// TIA Portal project "PROYECTO_FINALll" (V19)

(* hardware
DEVICE "PC-System_2"  SIMATIC PC station
   slot 0: "PC station"  Rail  SIMATIC PC-Station  V1.0
      slot 125: "Stationmanager"  Station_Manager  V6.0.4
   slot 1: "HMI_RT_1"  WinCC RT Advanced  6AV2 104-0xxxx-xxxx  17.0.0.0
      slot 33792: "Computer interface"  Host interface
   slot 2: "IE general_1"  IE General  IE_CP  V8.2.0
      slot 1: "PROFINET interface"  IEGeneral.Interface.8.2.0
DEVICE "S7-1200 station_2"  S7-1200 Station
   slot 0: "Rack_0"  S7-1200 Rack  Rack  V1.0
   slot 1: "PLC_2"  CPU 1212C AC/DC/Rly  6ES7 212-1BE40-0XB0  V4.5
   slot 101: "CM 1243-5"  CM 1243-5  6GK7 243-5DX30-0XE0  V1.3
DEVICE "GSD device_1"  GSD.Device
   slot 0: "Rack_0"  Rail
*)

// ===== PLC "PLC_2"  CPU 1212C AC/DC/Rly =====

VAR_GLOBAL   // PLC tag table "Default tag table"
   "Tag_1" AT %IW68 : Int;
   "Tag_2" AT %IW70 : Int;
   "Tag_3" AT %IW72 : Word;
   "Tag_4" AT %IW74 : Int;
   "Tag_5" AT %IW76 : Int;
   "Tag_6" AT %IW78 : Int;
END_VAR

DATA_BLOCK "Data"   // DB1
{ S7_Optimized_Access := 'TRUE' }
VERSION : 0.1
   VAR
      TEMP_A : Real;
      TEMP_M : Real;
      IRRADIANCIA : Real;
      SOILING : Real;
      VOLT_MED : Real;
      CORRIENTE_MED : Real;
      VDC : Real;
      IDC : Real;
      PAC : Real;
      PR : Real;
      YF : Real;
      EAC : Real;
      PERD_SUCIEDAD : Real;
      PERD_TEMP : Real;
      "ON/OFF" : Bool;
      DEFAULT : Bool;
   END_VAR
BEGIN
END_DATA_BLOCK

DATA_BLOCK "V_AMBIENTALES_DB"   // DB2
{ S7_Optimized_Access := 'TRUE' }
VERSION : 0.1
// stored: InstanceOfName V_AMBIENTALES
"V_AMBIENTALES"
BEGIN
END_DATA_BLOCK

DATA_BLOCK "Block_1_DB"   // DB3
{ S7_Optimized_Access := 'TRUE' }
VERSION : 0.1
// stored: InstanceOfName Block_1
"Block_1"
BEGIN
END_DATA_BLOCK

DATA_BLOCK "Block_1_DB_1"   // DB4
{ S7_Optimized_Access := 'TRUE' }
VERSION : 0.1
// stored: InstanceOfName Block_1
"Block_1"
BEGIN
END_DATA_BLOCK

FUNCTION_BLOCK "V_AMBIENTALES"   // FB1, LAD
{ S7_Optimized_Access := 'TRUE' }
VERSION : 0.1
   VAR_OUTPUT
      TEMP_M : Real;
      TEMP_A : Real;
      IRRADIANCIA : Real;
      SUCIEDAD : Real;
      VOLTAJE : Real;
      CORRIENTE : Real;
   END_VAR
   VAR_TEMP
      Temp_1 : Real;
      Temp_2 : Real;
      Temp_3 : Real;
      Temp_4 : Real;
      Temp_5 : Real;
      Temp_6 : Real;
   END_VAR
BEGIN

REGION Network 1: TEMPERATURA DEL MODULO
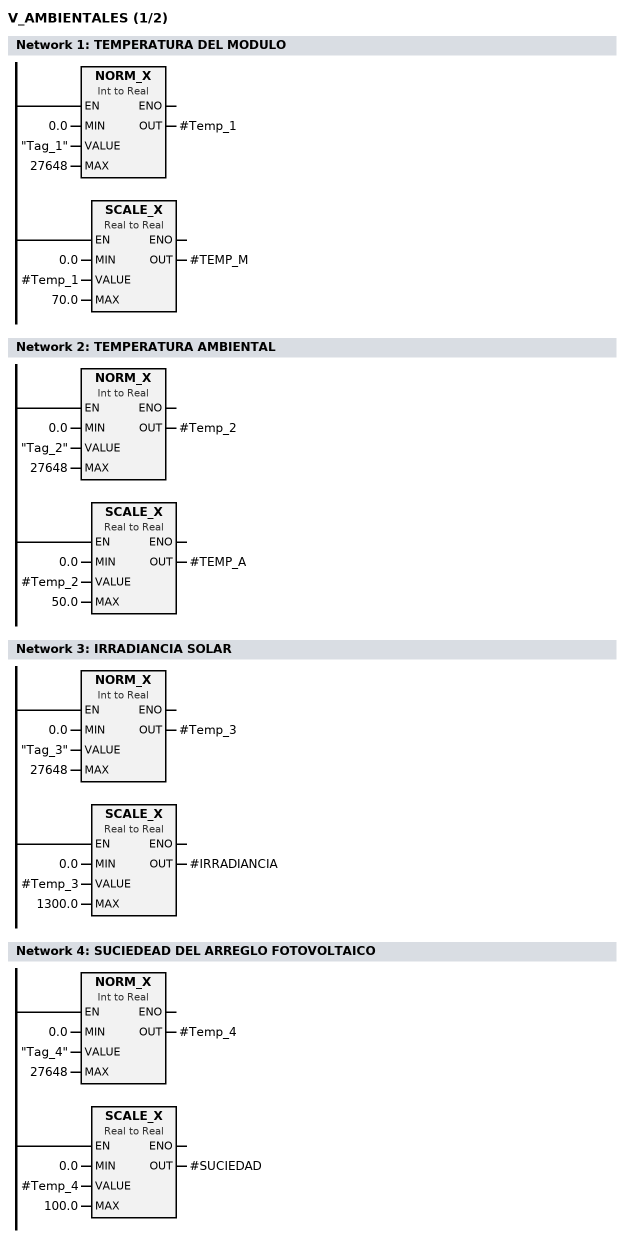
   RUNG wire#powerrail
      { S7_Templates := "[SrcType := Int, DestType := Real]" } Normalize(min := 0.0, value := "Tag_1", max := 27648, out => #Temp_1)
   END_RUNG
   RUNG wire#powerrail
      { S7_Templates := "[SrcType := Real, DestType := Real]" } Scale(min := 0.0, value := #Temp_1, max := 70.0, out => #TEMP_M)
   END_RUNG
   // the same network as SCL:
   #Temp_1 := NORM_X(MIN := 0.0, VALUE := "Tag_1", MAX := 27648);
   #TEMP_M := SCALE_X(MIN := 0.0, VALUE := #Temp_1, MAX := 70.0);
END_REGION

REGION Network 2: TEMPERATURA AMBIENTAL
   RUNG wire#powerrail
      { S7_Templates := "[SrcType := Int, DestType := Real]" } Normalize(min := 0.0, value := "Tag_2", max := 27648, out => #Temp_2)
   END_RUNG
   RUNG wire#powerrail
      { S7_Templates := "[SrcType := Real, DestType := Real]" } Scale(min := 0.0, value := #Temp_2, max := 50.0, out => #TEMP_A)
   END_RUNG
   // the same network as SCL:
   #Temp_2 := NORM_X(MIN := 0.0, VALUE := "Tag_2", MAX := 27648);
   #TEMP_A := SCALE_X(MIN := 0.0, VALUE := #Temp_2, MAX := 50.0);
END_REGION

REGION Network 3: IRRADIANCIA SOLAR
   RUNG wire#powerrail
      { S7_Templates := "[SrcType := Int, DestType := Real]" } Normalize(min := 0.0, value := "Tag_3", max := 27648, out => #Temp_3)
   END_RUNG
   RUNG wire#powerrail
      { S7_Templates := "[SrcType := Real, DestType := Real]" } Scale(min := 0.0, value := #Temp_3, max := 1300.0, out => #IRRADIANCIA)
   END_RUNG
   // the same network as SCL:
   #Temp_3 := NORM_X(MIN := 0.0, VALUE := "Tag_3", MAX := 27648);
   #IRRADIANCIA := SCALE_X(MIN := 0.0, VALUE := #Temp_3, MAX := 1300.0);
END_REGION

REGION Network 4: SUCIEDEAD DEL ARREGLO FOTOVOLTAICO
   RUNG wire#powerrail
      { S7_Templates := "[SrcType := Int, DestType := Real]" } Normalize(min := 0.0, value := "Tag_4", max := 27648, out => #Temp_4)
   END_RUNG
   RUNG wire#powerrail
      { S7_Templates := "[SrcType := Real, DestType := Real]" } Scale(min := 0.0, value := #Temp_4, max := 100.0, out => #SUCIEDAD)
   END_RUNG
   // the same network as SCL:
   #Temp_4 := NORM_X(MIN := 0.0, VALUE := "Tag_4", MAX := 27648);
   #SUCIEDAD := SCALE_X(MIN := 0.0, VALUE := #Temp_4, MAX := 100.0);
END_REGION

REGION Network 5: VOLTAJE DC
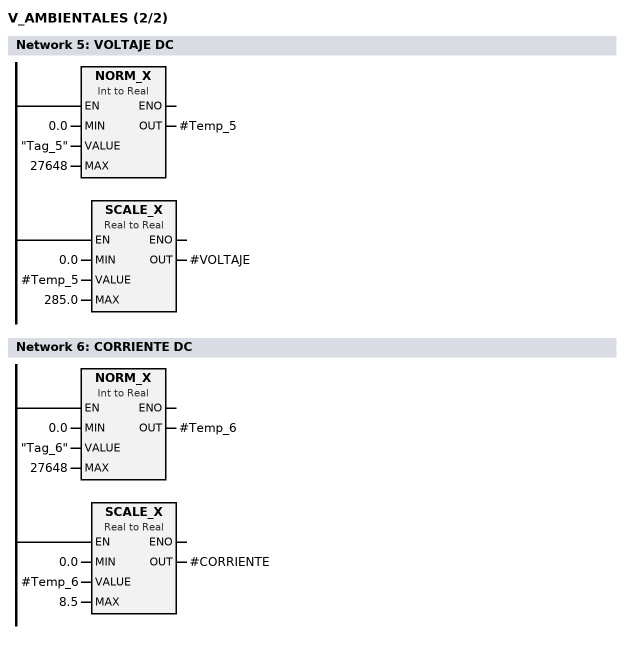
   RUNG wire#powerrail
      { S7_Templates := "[SrcType := Int, DestType := Real]" } Normalize(min := 0.0, value := "Tag_5", max := 27648, out => #Temp_5)
   END_RUNG
   RUNG wire#powerrail
      { S7_Templates := "[SrcType := Real, DestType := Real]" } Scale(min := 0.0, value := #Temp_5, max := 285.0, out => #VOLTAJE)
   END_RUNG
   // the same network as SCL:
   #Temp_5 := NORM_X(MIN := 0.0, VALUE := "Tag_5", MAX := 27648);
   #VOLTAJE := SCALE_X(MIN := 0.0, VALUE := #Temp_5, MAX := 285.0);
END_REGION

REGION Network 6: CORRIENTE DC
   RUNG wire#powerrail
      { S7_Templates := "[SrcType := Int, DestType := Real]" } Normalize(min := 0.0, value := "Tag_6", max := 27648, out => #Temp_6)
   END_RUNG
   RUNG wire#powerrail
      { S7_Templates := "[SrcType := Real, DestType := Real]" } Scale(min := 0.0, value := #Temp_6, max := 8.5, out => #CORRIENTE)
   END_RUNG
   // the same network as SCL:
   #Temp_6 := NORM_X(MIN := 0.0, VALUE := "Tag_6", MAX := 27648);
   #CORRIENTE := SCALE_X(MIN := 0.0, VALUE := #Temp_6, MAX := 8.5);
END_REGION
END_FUNCTION_BLOCK

FUNCTION_BLOCK "CALCULOS"   // FB2, LAD
{ S7_Optimized_Access := 'TRUE' }
VERSION : 0.1
   VAR_OUTPUT
      VOLTAJE_DC : Real;
   END_VAR
   VAR_TEMP
      TEMP_1 : Real;
      TEMP_2 : Real;
   END_VAR
BEGIN

REGION Network 1
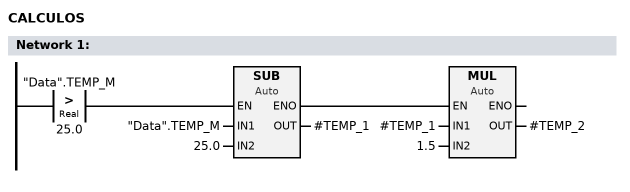
   RUNG wire#powerrail
      { S7_Templates := "SrcType := Real" } GT_Contact(in1 := "Data".TEMP_M, in2 := 25.0)
      Sub(in1 := "Data".TEMP_M, in2 := 25.0, out => #TEMP_1)
      Mul(in1 := #TEMP_1, in2 := 1.5, out => #TEMP_2)
   END_RUNG
   // the same network as SCL:
   IF "Data".TEMP_M > 25.0 THEN
       #TEMP_1 := "Data".TEMP_M - 25.0;
       #TEMP_2 := #TEMP_1 * 1.5;
   END_IF;
END_REGION
END_FUNCTION_BLOCK

FUNCTION_BLOCK "Block_1"   // FB3, SCL
{ S7_Optimized_Access := 'TRUE' }
VERSION : 0.1
   VAR_INPUT
      G_POA : Real;
      Tmod : Real;
      SR : Real;
      dt_s : Real;
      Enable : Bool;
      ResetDaily : Bool;
   END_VAR
   VAR_OUTPUT
      Vdc : Real;
      Idc : Real;
      Pac : Real;
      Eac : Real;
      Hpoa : Real;
      PR : Real;
      Yf : Real;
      Loss_soil : Real;
      Loss_therm : Real;
   END_VAR
   VAR
      P0_kw : Real := 2.25;
      Vdc_ref : Real := 282.0;
      Pac_max : Real := 2.0;
      eta_inv : Real := 0.96;
      gammaP : Real := 0.004;
      betaV : Real := 0.0035;
   END_VAR
   VAR_TEMP
      Geff : Real;
      Pdc : Real;
      tempFacP : Real;
      tempFacV : Real;
   END_VAR
BEGIN



   // Reset diario (por botón o por reloj)
   IF #ResetDaily THEN
       #Eac := 0.0;
       #Hpoa := 0.0;
   END_IF;

   IF NOT #Enable THEN
       // Si está deshabilitado, puedes congelar o poner en cero
       #Pac := 0.0;
       #Idc := 0.0;
       // Vdc lo puedes mantener o llevar a 0
       // Vdc := 0.0;
       #PR := 0.0;
       #Yf := #Eac / #P0_kw; // opcional
       RETURN;
   END_IF;

   // ---- Normalización y límites de SR ----
   // Si SR viene como porcentaje (0..100), lo convertimos a 0..1
   IF #SR > 1.5 THEN
       #SR := #SR / 100.0;
   END_IF;

   // Limitar SR a 0..1
   IF #SR < 0.0 THEN
       #SR := 0.0;
   ELSIF #SR > 1.0 THEN
       #SR := 1.0;
   END_IF;

   // ---- Pérdida por suciedad (%) ----
   #Loss_soil := 100.0 * (1.0 - #SR);

   // ---- Irradiancia efectiva (W/m²) ----
   IF #G_POA < 0.0 THEN
       #Geff := 0.0;
   ELSE
       #Geff := #G_POA * #SR;
   END_IF;

   // Factor térmico potencia (evitar que se haga >1.2 o negativo extremo)
   #tempFacP := 1.0 - #gammaP * (#Tmod - 25.0);
   IF #tempFacP < 0.0 THEN
       #tempFacP := 0.0;
   END_IF;

   // Pérdida térmica (solo si Tmod > 25)
   IF #Tmod > 25.0 THEN
       #Loss_therm := 100.0 * #gammaP * (#Tmod - 25.0);
   ELSE
       #Loss_therm := 0.0;
   END_IF;

   // Potencia DC (kW)
   #Pdc := #P0_kw * (#Geff / 1000.0) * #tempFacP;
   IF #Pdc < 0.0 THEN
       #Pdc := 0.0;
   END_IF;

   // Modelo de Vdc por temperatura
   #tempFacV := 1.0 - #betaV * (#Tmod - 25.0);
   IF #tempFacV < 0.2 THEN
       #tempFacV := 0.2;
   END_IF; // evita valores absurdos
   #Vdc := #Vdc_ref * #tempFacV;
   IF #Vdc < 50.0 THEN
       #Vdc := 50.0;
   END_IF;

   // Corriente DC (A)
   IF #Vdc > 0.0 THEN
       #Idc := (#Pdc * 1000.0) / #Vdc;
   ELSE
       #Idc := 0.0;
   END_IF;

   // Potencia AC (kW) + clipping
   #Pac := #eta_inv * #Pdc;
   IF #Pac > #Pac_max THEN
       #Pac := #Pac_max;
   END_IF;
   IF #Pac < 0.0 THEN
       #Pac := 0.0;
   END_IF;

   // Integraciones
   // Eac (kWh)
   #Eac := #Eac + (#Pac * #dt_s / 3600.0);

   // Hpoa (kWh/m²) desde G_POA (no Geff)
   #Hpoa := #Hpoa + (#G_POA * #dt_s / 3600000.0);

   // Rendimiento
   #Yf := #Eac / #P0_kw;

   // PR (%)
   IF #Hpoa > 0.01 THEN
       #PR := 100.0 * #Eac / (#P0_kw * #Hpoa);
   ELSE
       #PR := 0.0;
   END_IF;
END_FUNCTION_BLOCK

ORGANIZATION_BLOCK "Main"   // OB1, LAD, ProgramCycle
TITLE = "Main Program Sweep (Cycle)"
{ S7_Optimized_Access := 'TRUE' }
VERSION : 0.1
   VAR_INPUT
      Initial_Call : Bool;   // Initial call of this OB
      Remanence : Bool;   // =True, if remanent data are available
   END_VAR
BEGIN

REGION Network 1
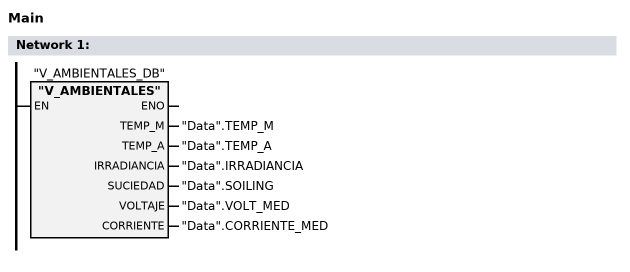
   RUNG wire#powerrail
      "V_AMBIENTALES_DB"(TEMP_M => "Data".TEMP_M, TEMP_A => "Data".TEMP_A, IRRADIANCIA => "Data".IRRADIANCIA, SUCIEDAD => "Data".SOILING, VOLTAJE => "Data".VOLT_MED, CORRIENTE => "Data".CORRIENTE_MED)
   END_RUNG
   // the same network as SCL:
   "V_AMBIENTALES_DB"(TEMP_M => "Data".TEMP_M,   // "V_AMBIENTALES"
                      TEMP_A => "Data".TEMP_A,
                      IRRADIANCIA => "Data".IRRADIANCIA,
                      SUCIEDAD => "Data".SOILING,
                      VOLTAJE => "Data".VOLT_MED,
                      CORRIENTE => "Data".CORRIENTE_MED);
END_REGION
END_ORGANIZATION_BLOCK

ORGANIZATION_BLOCK "CyclicInterrupt"   // OB30, LAD, CyclicInterrupt
{ S7_Optimized_Access := 'TRUE' }
VERSION : 0.1
   VAR_INPUT
      Initial_Call : Bool;   // Initial call of this OB
      Event_Count : Int;   // Events discarded
   END_VAR
   VAR_TEMP   // added for the SCL form of the ladder/FBD networks
      _w1 : Bool;
   END_VAR
BEGIN

REGION Network 1
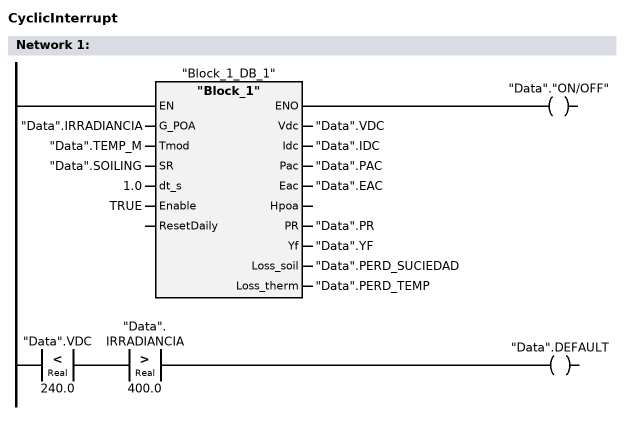
   RUNG wire#powerrail
      "Block_1_DB_1"(G_POA := "Data".IRRADIANCIA, Tmod := "Data".TEMP_M, SR := "Data".SOILING, dt_s := 1.0, Enable := TRUE, ResetDaily :=, Vdc => "Data".VDC, Idc => "Data".IDC, Pac => "Data".PAC, Eac => "Data".EAC, Hpoa =>, PR => "Data".PR, Yf => "Data".YF, Loss_soil => "Data".PERD_SUCIEDAD, Loss_therm => "Data".PERD_TEMP)
      Coil( "Data"."ON/OFF" )
   END_RUNG
   RUNG wire#powerrail
      { S7_Templates := "SrcType := Real" } LT_Contact(in1 := "Data".VDC, in2 := 240.0)
      { S7_Templates := "SrcType := Real" } GT_Contact(in1 := "Data".IRRADIANCIA, in2 := 400.0)
      Coil( "Data".DEFAULT )
   END_RUNG
   // the same network as SCL:
   "Block_1_DB_1"(G_POA := "Data".IRRADIANCIA,   // "Block_1"
                  Tmod := "Data".TEMP_M,
                  SR := "Data".SOILING,
                  dt_s := 1.0,
                  Enable := TRUE,
                  Vdc => "Data".VDC,
                  Idc => "Data".IDC,
                  Pac => "Data".PAC,
                  Eac => "Data".EAC,
                  PR => "Data".PR,
                  Yf => "Data".YF,
                  Loss_soil => "Data".PERD_SUCIEDAD,
                  Loss_therm => "Data".PERD_TEMP,
                  ENO => #_w1);
   "Data"."ON/OFF" := #_w1;
   "Data".DEFAULT := ("Data".VDC < 240.0) AND ("Data".IRRADIANCIA > 400.0);
END_REGION
END_ORGANIZATION_BLOCK

(* ===== HMI "HMI_RT_1" =====
system functions are stored by id; their names below are inferred from use
connection "HMI_Connection_1": ETHERNET, S7_1200_OMS
connection "HMI_Connection_2": ETHERNET, S7_1200_OMS

HMI tags "Default tag table"
   "Data_TEMP_M" : Real = PLC Data.TEMP_M, 100 ms
   "Data_IRRADIANCIA" : Real = PLC Data.IRRADIANCIA, 1 s
   "Data_TEMP_A" : Real = PLC Data.TEMP_A, 100 ms
   "Data_SOILING" : Real = PLC Data.SOILING, 100 ms
   "Data_VOLT_DC" : Real = PLC Data.VOLT_MED, 100 ms
   "Data_CORRIENT_DC" : Real = PLC Data.CORRIENTE_MED, 100 ms
   "Data_VDC" : Real = PLC Data.VDC, 100 ms
   "Data_IDC" : Real = PLC Data.IDC, 100 ms
   "Data_PAC" : Real = PLC Data.PAC, 1 s
   "Data_EAC" : Real = PLC Data.EAC, 100 ms
   "Data_PR" : Real = PLC Data.PR, 100 ms
   "Data_YF" : Real = PLC Data.YF, 100 ms
   "Data_PERD_SUCIEDAD" : Real = PLC Data.PERD_SUCIEDAD, 100 ms
   "Data_PERD_TEMP" : Real = PLC Data.PERD_TEMP, 100 ms
   "Data_ON/OFF" : Bool = PLC Data.ON/OFF, 100 ms
   "Data_DEFAULT" : Bool = PLC Data.DEFAULT, 100 ms

screen "Screen_1" 1024x768, template "Template_1"
   TextField "Text field_1" at 32,74 size 233x27; Text 'Irradiancia POA (W/m²)'
   TextField "Text field_2" at 347,23 size 305x36; Text 'Variables ambientales'
   TextField "Text field_4" at 341,73 size 292x27; Text 'Temperatura del módulo (°C)'
   TextField "Text field_5" at 710,72 size 269x27; Text 'Temperatura ambiente (°C)'
   IOField "I/O field_1" at 83,98 size 112x23; FormatPattern 9999
      ProcessValue <- "Data_IRRADIANCIA"
   IOField "I/O field_2" at 438,98 size 112x24; FormatPattern 9999.9
      ProcessValue <- "Data_TEMP_M"
   IOField "I/O field_3" at 805,97 size 112x25; FormatPattern 99999.9
      ProcessValue <- "Data_TEMP_A"
   TextField "Text field_6" at 38,136 size 278x27; Text 'Proporcion por suciedad (%)'
   IOField "I/O field_4" at 113,160 size 112x25; FormatPattern 999
      ProcessValue <- "Data_SOILING"
   TextField "Text field_7" at 362,207 size 278x36; Text 'Variables electricas'
   TextField "Text field_8" at 70,263 size 165x27; Text 'Voltaje DC (Vdc)'
   TextField "Text field_10" at 409,262 size 184x27; Text 'Corriente DC (Idc)'
   IOField "I/O field_5" at 90,286 size 112x26; FormatPattern 999.9
      ProcessValue <- "Data_VDC"
   IOField "I/O field_6" at 442,285 size 112x27; FormatPattern 99.9
      ProcessValue <- "Data_IDC"
   IOField "I/O field_7" at 801,286 size 112x25; FormatPattern 9999.9
      ProcessValue <- "Data_PAC"
   TextField "Text field_11" at 20,336 size 288x27; Text 'Energía AC acumulada (kWh)'
   IOField "I/O field_8" at 89,362 size 112x24; FormatPattern 9999.9
      ProcessValue <- "Data_EAC"
   TextField "Text field_12" at 780,260 size 176x27; Text 'Potencia AC (kW)'
   TextField "Text field_13" at 404,336 size 194x25; Text 'Estado del inversor'
   TextField "Text field_14" at 414,364 size 76x27; Text 'ON/OFF'
   TextField "Text field_16" at 530,363 size 57x27; Text 'FAULT'
   GraphicIOField "PlotLight_Round_GN" at 429,389 size 34x34; PictureOff "PilotLight_Round_GN_Off_256c"; PictureOn "PilotLight_Round_GN_On_256c"
      ProcessValue <- "Data_ON/OFF"
   GraphicIOField "PlotLight_Round_RN" at 541,389 size 34x35; PictureOff "PilotLight_Round_RN_Off_256c"; PictureOn "PilotLight_Round_RN_On_256c"
      ProcessValue <- "Data_DEFAULT"
   TextField "Text field_17" at 335,454 size 343x36; Text 'Variables de rendimiento'
   TextField "Text field_18" at 33,504 size 237x27; Text 'Factor de potencia (FP)'
   TextField "Text field_19" at 391,504 size 230x27; Text 'Performance Ratio (%)'
   TextField "Text field_20" at 663,503 size 343x27; Text 'Rendimiento específico (kWh/kHp)'
   IOField "I/O field_10" at 88,528 size 112x25; FormatPattern 999999999999
   IOField "I/O field_11" at 450,529 size 112x24; FormatPattern 99.99
      ProcessValue <- "Data_PR"
   IOField "I/O field_12" at 788,529 size 112x25; FormatPattern 99.99
      ProcessValue <- "Data_YF"
   TextField "Text field_21" at 432,586 size 121x36; Text 'Perdidas'
   IOField "I/O field_13" at 190,660 size 112x23; FormatPattern 99.99
      ProcessValue <- "Data_PERD_TEMP"
   TextField "Text field_22" at 139,634 size 222x27; Text 'Pérdidas térmicas (%)'
   TextField "Text field_23" at 612,634 size 261x27; Text 'Pérdidas por suciedad (%)'
   IOField "I/O field_14" at 681,660 size 112x24; FormatPattern 99.99
      ProcessValue <- "Data_PERD_SUCIEDAD"
   Button "Button_2" at 196,99 size 42x22; TextOff 'Gráf'
      on Press: ActivateScreen("Screen_4", 0)
   Button "Button_3" at 552,98 size 42x22; TextOff 'Gráf'
      on Press: ActivateScreen("Screen_5", 0)
   Button "Button_4" at 919,97 size 42x22; TextOff 'Gráf'
      on Press: ActivateScreen("Screen_6", 0)
   Button "Button_5" at 204,287 size 42x22; TextOff 'Gráf'
      on Press: ActivateScreen("Screen_7", 0)
   Button "Button_6" at 556,286 size 42x22; TextOff 'Gráf'
      on Press: ActivateScreen("Screen_8", 0)
   Button "Button_7" at 914,287 size 42x22; TextOff 'Gráf'
      on Press: ActivateScreen("Screen_9", 0)

Template "Template_1" 1024x768
   Button "Template_Button_1" at 10,714 size 104x34; TextOff 'SALIR'
      on Press: StopRuntime(0)
   Button "Template_Button_2" at 789,698 size 46x46; TextOff 'P1'
      on Press: ActivateScreen("Screen_1", 0)
   Button "Template_Button_3" at 863,698 size 46x46; TextOff 'P2'
      on Press: ActivateScreen("Screen_2", 0)
   Button "Template_Button_4" at 937,698 size 46x46; TextOff 'P3'
      on Press: ActivateScreen("Screen_3", 0)

screen "Screen_2" 1024x768, template "Template_1"
   TextField "Text field_1" at 268,26 size 473x39; Text 'Comparación POA vs. Potencia'
   TrendView "Trend view_1" at 16,80 size 989x589

screen "Screen_3" 1024x768, template "Template_1"
   TextField "Text field_1" at 332,23 size 340x39; Text 'ENERGIA ACOMULADA'
   TrendView "Trend view_1" at 15,89 size 988x580

screen "Screen_4" 1024x768, template "Template_2"
   TextField "Text field_1" at 338,25 size 366x39; Text 'IRRADIANCIA vs TIEMPO'
   TrendView "Trend view_1" at 15,89 size 988x580

Template "Template_2" 1024x768
   Button "Template_Button_1" at 10,714 size 104x34; TextOff 'VOLVER'
      on Press: ActivateScreen("Screen_1", 0)

screen "Screen_5" 1024x768, template "Template_2"
   TextField "Text field_1" at 311,25 size 359x39; Text 'T° MODULOS vs TIEMPO'
   TrendView "Trend view_1" at 15,89 size 988x580

screen "Screen_6" 1024x768, template "Template_2"
   TextField "Text field_1" at 333,25 size 363x39; Text 'T° AMBIENTE vs TIEMPO'
   TrendView "Trend view_1" at 15,89 size 988x580

screen "Screen_7" 1024x768, template "Template_2"
   TextField "Text field_1" at 342,26 size 329x39; Text 'VOLTAJE DC vs TIEMO'
   TrendView "Trend view_1" at 15,89 size 988x580

screen "Screen_8" 1024x768, template "Template_2"
   TextField "Text field_1" at 323,26 size 384x39; Text 'CORRIENTE DC vs TIEMPO'
   TrendView "Trend view_1" at 15,100 size 988x580

screen "Screen_9" 1024x768, template "Template_2"
   TextField "Text field_1" at 329,26 size 368x39; Text 'POTENCIA AC vs TIEMPO'
   TrendView "Trend view_1" at 15,89 size 988x580
*)